PROGRAM main
  VAR
    S1 AT %IX0.0  : BOOL; (* marcha, NA *)
    S0 AT %IX0.1  : BOOL; (* parada, NC: TRUE sin pulsar *)
    KM1 AT %QX0.0 : BOOL; (* línea *)
    KM2 AT %QX0.1 : BOOL; (* estrella *)
    KM3 AT %QX0.2 : BOOL; (* triángulo *)
    H1 AT %QX0.3  : BOOL; (* piloto en marcha *)
    ETAPA         : INT; (* 0 parado, 1 estrella, 2 pausa, 3 triángulo *)
    T_EST         : TON;
    T_PAU         : TON;
    FIN_EST       : BOOL;
    FIN_PAU       : BOOL;
    E0            : BOOL; (* ETAPA = 0 *)
    E1            : BOOL; (* ETAPA = 1 *)
    E2            : BOOL; (* ETAPA = 2 *)
    E3            : BOOL; (* ETAPA = 3 *)
  END_VAR

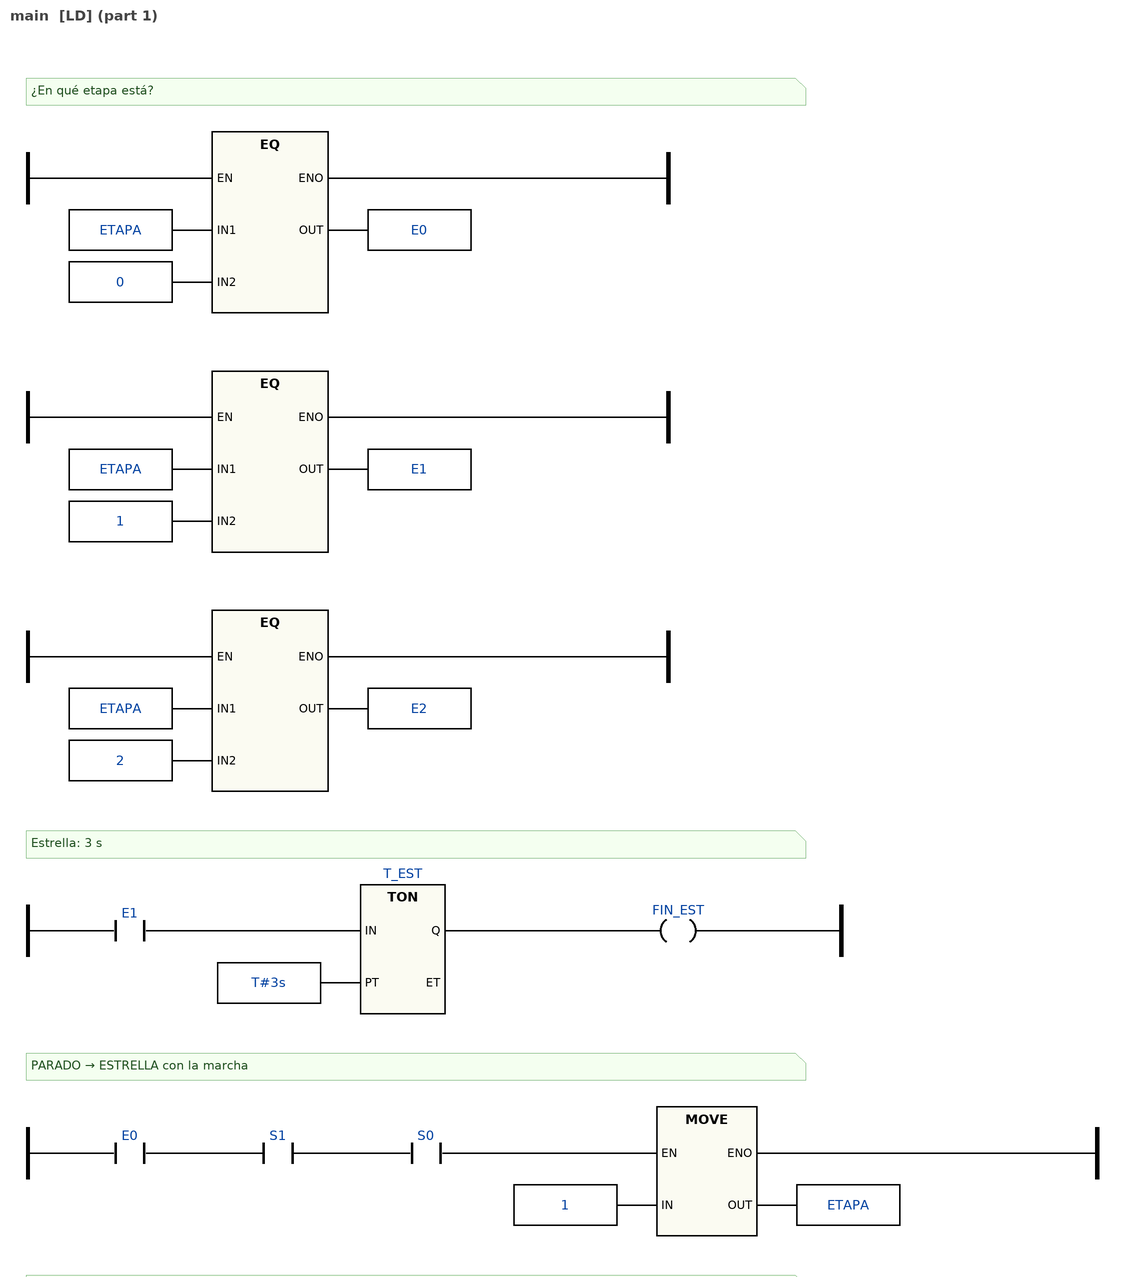
(* LD diagram, written out as Structured Text *)
(* ¿En qué etapa está? *)
E0 := ETAPA = 0;
E1 := ETAPA = 1;
E2 := ETAPA = 2;
(* Estrella: 3 s *)
T_EST(IN := E1, PT := T#3s);
FIN_EST := T_EST.Q;
(* PARADO → ESTRELLA con la marcha *)
IF E0 AND S1 AND S0 THEN ETAPA := 1; END_IF;
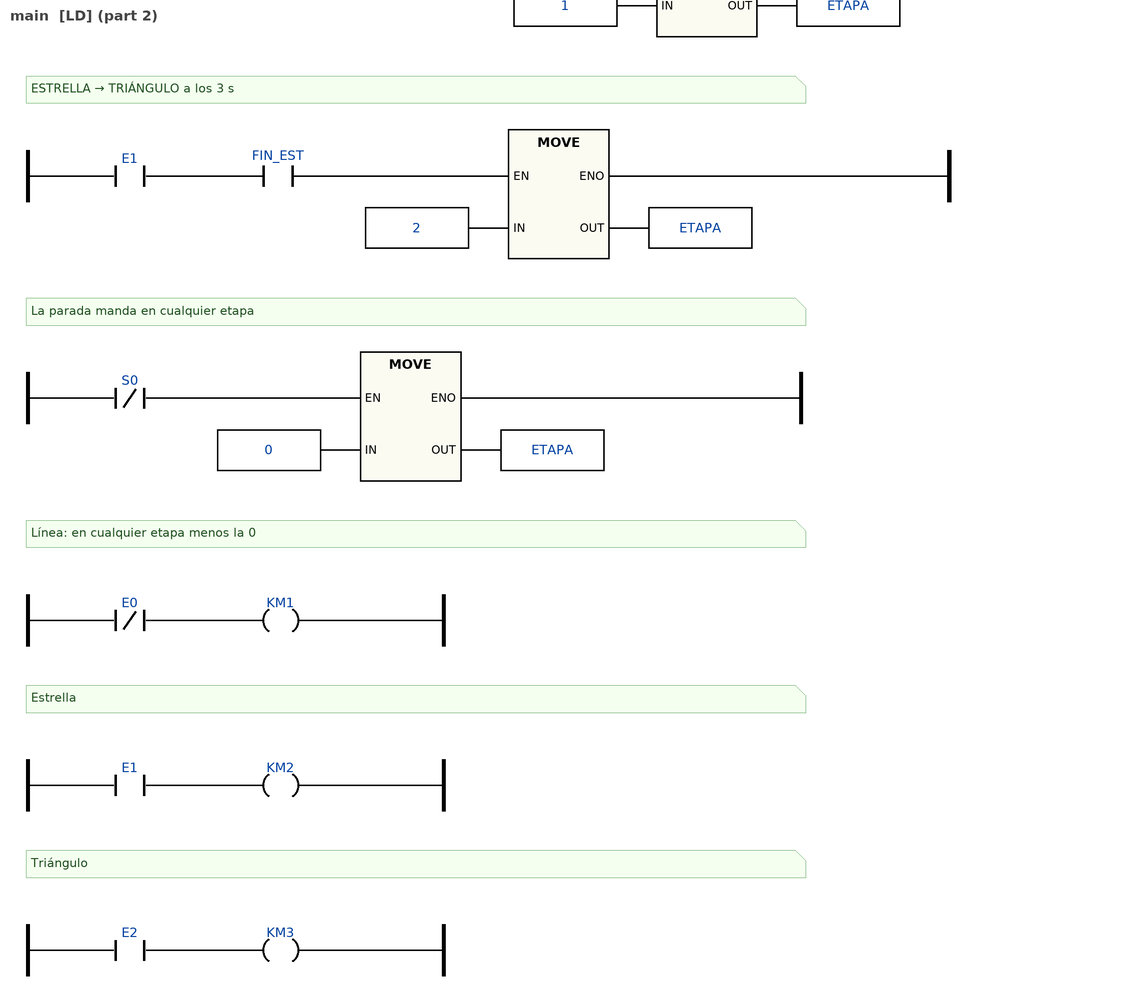
(* ESTRELLA → TRIÁNGULO a los 3 s *)
IF E1 AND FIN_EST THEN ETAPA := 2; END_IF;
(* La parada manda en cualquier etapa *)
IF NOT S0 THEN ETAPA := 0; END_IF;
(* Línea: en cualquier etapa menos la 0 *)
KM1 := NOT E0;
(* Estrella *)
KM2 := E1;
(* Triángulo *)
KM3 := E2;
END_PROGRAM
